(* IEC 61131-3 sources: codesys-to-s7/tests/corpus/C2S7-TYPE-RANGE/pos, 1 file *)

(* ---- input.st ---- *)
FUNCTION_BLOCK FB_Case
VAR
    x : INT(0..100);
END_VAR
x := 5;
END_FUNCTION_BLOCK
